// TIA Portal V21 export
// export: Created 2026-11-22T04:06:07.4620333Z, ExportSetting WithDefaults, DisplayName Totally Integrated Automation Portal, DisplayVersion V21 Update 3, DisplayName STEP 7 Professional, DisplayVersion V21 Update 3, DisplayName STEP 7 Safety, DisplayVersion V21, DisplayName Tech WebApplication, DisplayVersion V21, DisplayName WinCC Basic/Comfort/Advanced, DisplayVersion V21 Update 3, DisplayName WinCC Unified, DisplayVersion V21 Update 3
VBScript "C5_ToggleSlideIn"  Type=Sub
  ShowSlideInScreen "Slide-in screen top", hmiToggle
